Fanuc KAREL source: kt00008.KL

-- PROVISIONAL review KL for V940-1; original PC SHA256 b444f33920c8672285e28de1c2f26d4a481263bf0300dae77cf650c8a7d003c7
-- Incomplete behavior may be omitted. Consult companion uncertainty JSON. Do not deploy.
PROGRAM KT00008
%NOLOCKGROUP
VAR
  I1 : INTEGER
  OUT : REAL
-- UNRESOLVED_DECL H2 type=002017
BEGIN
  -- V9_ZERO_TABLE_METADATA_HINT layout=0001; no indexed target words; source/name/runtime held
  -- UNRESOLVED_PC offsets 5-16; opcodes 2E,23
  -- UNRESOLVED_PC offsets 21-35; opcodes 2E,22,9D,33,B4
  -- UNRESOLVED_PC offsets 40-63; opcodes 21,22,9D,33,B3,52,64,23
  -- UNRESOLVED_PC offsets 68-72; opcodes 7F
END KT00008
